(* IEC 61131-3 sources: kns-port-domestic/targets/astra/src/POUs/Log/FB_DeviceAudit, 2 files *)

(* ---- FB_DeviceAudit.decl.st ---- *)
// Назначение: аудит режимов устройств перечня (GVL_Log.fbDeviceAudit, MainTask после PRG_Devices… вызывает
//             PRG_Station): смена Mode устройства — событие станции 101018 со значением dev_no · 10 + режим
//             (E_DeviceMode). Первый вызов запоминает режимы без событий (режимы после старта — из retain).
// Автор:      kr0nsch
// Версия:     0.1.1
// Документ:   docs/DESIGN.md, раздел 9.3; docs/04_algorithms.md, раздел 16
FUNCTION_BLOCK FB_DeviceAudit
VAR_INPUT
    aitfDevice : ARRAY[1..GVL_DeviceList.DEVICE_COUNT] OF PL.I_Device;   // GVL_DeviceList.aitfDevice
    auiDevNo   : ARRAY[1..GVL_DeviceList.DEVICE_COUNT] OF UINT;          // GVL_DeviceList.auiDevNo
    itfEvents  : I_StationEventSink;                                     // журнал; 0 — без событий
END_VAR
VAR_OUTPUT
    udiChanges : UDINT;             // замечено смен режима с запуска
END_VAR
VAR
    aeModePrev : ARRAY[1..GVL_DeviceList.DEVICE_COUNT] OF PL.E_DeviceMode;   // режим прошлого вызова
    axKnown    : ARRAY[1..GVL_DeviceList.DEVICE_COUNT] OF BOOL;             // режим устройства уже запомнен
    uiI        : UINT;              // индекс устройства
    eMode      : PL.E_DeviceMode;   // режим этого вызова
    itfDev     : PL.I_Device;       // устройство
END_VAR

(* ---- FB_DeviceAudit.impl.st ---- *)
FOR uiI := 1 TO GVL_DeviceList.DEVICE_COUNT DO
    itfDev := aitfDevice[uiI];
    IF itfDev <> 0 THEN
        eMode := itfDev.Mode;
        IF axKnown[uiI] AND eMode <> aeModePrev[uiI] THEN
            udiChanges := udiChanges + 1;
            IF itfEvents <> 0 THEN
                // в UDINT: dev_no до 9999 (API 20.1) · 10 не помещается в UINT
                itfEvents.LogEvent(eEvent := E_StationEvent.DeviceModeChanged,
                                   rValue := UDINT_TO_REAL(UINT_TO_UDINT(auiDevNo[uiI])
                                                           * UINT_TO_UDINT(GVL_Const.LOG_DEV_MODE_SCALE)
                                                           + TO_UDINT(eMode)));
            END_IF
        END_IF
        aeModePrev[uiI] := eMode;
        axKnown[uiI] := TRUE;
    END_IF
END_FOR
